(* IEC 61131-3 sources: JingjiangArm/moonboxpro_arm_8.4/Application/Application/数据类型/通讯协议/云影/只写内容/附属内容, 6 files *)

(* ---- StSts_GrpFlag.st ---- *)
(*@CES
Name=StSts_GrpFlag
Type=Gvl
TypeGuid=2db5746d-d284-4425-9f7f-2663a34b0ebc
Guid=84c3180d-bd4c-42e6-a1a9-68017632a9f9
HasDeclaration=True
HasImplementation=False
*)
{DECLARATION}
{attribute 'pack_mode' := '1'}
TYPE StSts_GrpFlag :(*2025.7.3.175755总16字节+8预留字节*)
STRUCT
	xCutterOnTop_Uw								: BIT;(* TRUE=放料上裁 *)
	xCutterOnTop_Rw								: BIT;(* TRUE=放料上裁 *)
	xFlag_Stop									: BIT;(* 停机标志/第1次从当前速度降到空转速度，抬所有色组胶辊/牵引速度到0时抬牵引胶辊，第2次按下则将色组从空转停到0速度 *)
	xFlag_PreStart								: BIT;(* 预启动标志/从停机状态按(预)启动置位标志 色组速度达到空转速度清xFlag_PreStart标志,置位xFlag_Ink标志;当xFlag_Print标志有效后 *)
	xFlag_Ink									: BIT;(* 匀墨标志/>20m/min不能联动 *)
	xFlag_InkAccing								: BIT;(* 匀墨加速中<指0~10m/min那个加速过程> *)
	xFlag_Tension								: BIT;(* 张力投入标志/张力投入有效时收放料变频开始起作用/收放料就位后按印刷按钮,牵引压辊合压/xFlag_Print有效时张力投入不处理 *)
	xFlag_TensionDone							: BIT;(* 张力ok，可以投入印刷 *)
	xFlag_Print									: BIT;(* 张力拉料标志有效时，按联动或印刷按钮 先压收牵(延时2s)再压放牵 印刷标志/印刷色组根据联动标志按用户指定的压辊顺序逐一延时压胶辊/胶辊压合完毕后才可置该标志有效 *)
	xFlag_Estop									: BIT;(* 急停标志/和停机一样要减速到0，只不过减速时间是急停时间 *)
	xFlag_AutoAcc								: BIT;(* 自动加速 *)
	xFlag_AutoDec								: BIT;(* 自动减速 *)
	xFlag_ManuAcc								: BIT;(* 手动加速 *)
	xFlag_ManuDec								: BIT;(* 手动减速 *)
	xFlag_Accing								: BIT;(* 加速中 *)
	xFlag_Decing								: BIT;(* 减速中 *)
	xFlag_EStoping								: BIT;(* 正在急停中 *)
	xFlag_Stoping								: BIT;(* 停机中 *)
	xFlag_GotoInking							: BIT;(* 转到匀墨 *)
	xFlag_InPressing							: BIT;(* 顺序压辊中 *)
	xFlag_RollerPressDone						: BIT;(* 压辊处理完成 *)
	xFlag_InchRun								: BIT;(* 至少有1色处于单运行 *)
	xFlag_AllInchRun							: BIT;(* 整机单运行标志 *)
	xFlag_AllPress								: BIT;(* 全体合压 *)
	xFlag_AllUnpress							: BIT;(* 全体离压 *)
	xFlag_RollerPressAtLeast1					: BIT;(* 至少1色色组合压 *)
	xFlag_PrnLen_Alarm_A						: BIT;
	xFlag_PrnLen_Alarm_B						: BIT;
	xFlag_PrnLen_Alarm_All						: BIT;
	xFlag_LinkageAxisAlarm						: BIT;(* 至少有1个联动轴发生报警 *)
	xFlag_TensionUnfinished						: BIT;(* 张力未完成 *)
	xFlag_VelTooHigh							: BIT;(* 速度过高 *)
	xFlag_PrestartTimeout						: BIT;(* 预启动超时标志 *)
	xFlag_KeepAlarming							: BIT;(* 维持报警*)
	xFlag_ArrivedToTargetVel					: BIT;(* 到达目标速度 *)
	xFlag_FilmAccDecDone						: BIT;(* 料膜加减速完成 *)
	xFlag_IfOf_Ink								: BIT;(*空转牵引联动标志*)
	xFlag_FastStoping							: BIT;
	xSlowStopTenEn								: BIT;(* 收放料慢速松料使能/TRUE *)
	xIsDebugMode_Machine						: BIT;(* 机器调试模式 *)
(*以上40bit*)
	xReflectSensorLoss_Uw						: BIT;(* 放料弧面信号丢失标志/FALSE *)
	xFilmTouchRoller_Uw							: BIT;(*料膜接触到了辊子标志*)
	xSts_PreCutting_Uw							: BIT;(* 放料预备接料/FALSE *)
	xCutterOnTopFroDebug_Uw						: BIT;(* 放料上裁刀标志/用于调试/FALSE *)
	xCurAxisAFroDebug_Uw						: BIT;(* 放料预驱轴为A轴标志/用于调试/FALSE *)
	xAlarmBell_Uw								: BIT;(* 放料响铃常输出/用于控制定位写入响铃提示使用/FALSE *)
	xIsDebuging_DiaMeasure_Uw					: BIT;(* 放料卷径测量调试中/FALSE *)
	xCancelDebuging_DiaMeasure_Uw				: BIT;(* 放料取消卷径测量调试中/FALSE *)
	xEnCodeErr_Uw								: BIT;(* 放料编码器故障*)
	xEnCodeErr_Rw								: BIT;(* 收料编码器故障*)
	xAxisAForeward_Uw							: BIT;(* 放料A轴正转/FALSE *)
	xAxisBForeward_Uw							: BIT;(* 放料B轴正转/FALSE *)
	xFlag_DiamCalc_ing_Uw						: BIT;(* 放料卷径计算中 *)
	xFlag_DiamCalc_end_Uw						: BIT;(* 放料卷径计算完成 *)
	xFlag_DiamMeasure_end_Uw					: BIT;(* 放料卷径测量完成 *)
	xFlag_PreDrv_ing_Uw							: BIT;(* 放料预驱中... *)
	xFlag_PreDrv_end_Uw							: BIT;(* 放料预驱完成  *)
	xFlag_Cut_ing_Uw							: BIT;
	xFlag_Cut_end_Uw							: BIT;
	xFlag_VolDiamAlarm_Uw						: BIT;(* 卷径报警标志 *)
	xStationOnline_AxisA_Uw						: BIT;(* 放料a轴驱动器在线标志/2021.12.4.175524/hdp *)
	xStationOnline_AxisB_Uw						: BIT;(* 放料a轴驱动器在线标志/2021.12.4.175524/hdp *)
	xFlag_AutoMaticCutting_Uw					: BIT;(*2022.4.25.090246 自动裁切中标志*)
(*以上23bit*)
	xSts_PreCutting_Rw							: BIT;(* 收料预备接料 *)
	xCutterOnTopFroDebug_Rw						: BIT;(* 收料上裁刀标志/用于调试/FALSE *)
	xCurAxisAFroDebug_Rw						: BIT;(* 收料预驱轴为A轴标志/用于调试/FALSE *)
	x6InchFroDebug_Rw       					: BIT;(* 收料6寸标志/用于调试/FALSE*)
	xAlarmBell_Rw								: BIT;(* 收料响铃常输出/用于控制定位写入响铃提示使用/FALSE *)
	xAxisAForeward_Rw							: BIT;(* 收料A轴正转/FALSE *)
	xAxisBForeward_Rw							: BIT;(* 收料B轴正转/FALSE *)
	xFlag_6Inch_Rw								: BIT;(* 收料6寸标志/反之为3寸/FALSE *)
	xFlag_PreDrv_ing_Rw							: BIT;(* 收料预驱中... *)
	xFlag_PreDrv_end_Rw							: BIT;(* 收料预驱完成 *)
	xFlag_Cut_ing_Rw							: BIT;(* 收料裁切中 *)
	xFlag_Cut_end_Rw							: BIT;(* 收料裁切完成 *)
	xStationOnline_AxisA_Rw						: BIT;(* 收料a轴驱动器在线标志/2021.12.4.175524/hdp *)
	xStationOnline_AxisB_Rw						: BIT;(* 收料a轴驱动器在线标志/2021.12.4.175524/hdp *)
	xFlag_AutoMaticCutting_rw					: BIT;(*2022.4.25.090246 自动裁切中标志*)
(*以上15bit*)
	xStationOnline_If							: BIT;(* 放牵驱动器在线标志/2021.12.4.175524/hdp *)
	xRollerSts_If								: BIT;(* 放牵压辊/FALSE *)
	xRunEn_If									: BIT;(* 放牵运动使能/0/2021.11.18.201925 *)
	xInching_If									: BIT;(* 放牵单运行中/FALSE *)
	xStationOnline_Of							: BIT;(* 放牵驱动器在线标志/2021.12.4.175524/hdp *)
	xRollerSts_Of								: BIT;(* 放牵压辊/FALSE *)
	xRunEn_Of									: BIT;(* 放牵运动使能/0/2021.11.18.201925 *)
	xInching_Of									: BIT;(* 放牵单运行中/FALSE *)
(*以上8bit*)
	xSts_HorzPreRegister						: BIT;(*横向预套准状态*)
	xFlag_HorzPreRegister_All_end				: BIT;(*横向预套准全部完成*)
	xFlag_Home									: BIT;
	xFlag_Home_ing								: BIT;
	xFlag_Home_end								: BIT;
	xFlag_ConfirmPreRegHomePos					: BIT;(*2017-09-13 12:51:52| 确认预套准基准点*)
	xFlag_ConfirmPreRegHomePos_ing				: BIT;(*确认预套准基准点-ing*)
	xFlag_ConfirmPreRegHomePos_end				: BIT;(*确认预套准基准点-end*)
	xFlag_PreRegister							: BIT;
	xFlag_PreRegister_ing						: BIT;
	xFlag_PreRegister_end						: BIT;
	xFlag_PhaseRestore							: BIT;(*相位恢复*)
	xFlag_PhaseRestore_ing						: BIT;(*相位恢复-ing*)
	xFlag_PhaseRestore_end						: BIT;(*相位恢复-end*)
(*以上14bit*)
	xNetOffline_CENTRAL							: BIT;
	xAxisAlarm_CENTRAL							: BIT;
	xPosDeviationAlarm_CENTRAL					: BIT;
	xNetOffline_CENTRAL2						: BIT;
	xAxisAlarm_CENTRAL2							: BIT;
	xPosDeviationAlarm_CENTRAL2					: BIT;
	xNetOffline_IF								: BIT;
	xAxisAlarm_IF								: BIT;
	xPosDeviationAlarm_IF						: BIT;
	xNetOffline_OF								: BIT;
	xAxisAlarm_OF								: BIT;
	xPosDeviationAlarm_OF						: BIT;
	xNetOffline_UW_A							: BIT;
	xAxisAlarm_UW_A								: BIT;
	xPosDeviationAlarm_UW_A						: BIT;
	xNetOffline_UW_B							: BIT;
	xAxisAlarm_UW_B								: BIT;
	xPosDeviationAlarm_UW_B						: BIT;
	xNetOffline_RW_A							: BIT;
	xAxisAlarm_RW_A								: BIT;
	xPosDeviationAlarm_RW_A						: BIT;
	xNetOffline_RW_B							: BIT;
	xAxisAlarm_RW_B								: BIT;
	xPosDeviationAlarm_RW_B						: BIT;
	xPrintInching								: BIT;//整机点动
	xTapPosition_Breaking						: BIT;(*断料档位|*)
	xTapPosition_UniformInk						: BIT;(*匀墨档位|*)
	xTapPosition_Printing						: BIT;(*印刷档位|*)
(*以上28bit*)
////////////////////////////////////////////////////////////////////////////////////
(*截至这里，以上总共40+23+15+8+14+28=128BIT，占16BYTES，下面再预留8BYTE，用于放系只写标志*)
(*2025.9.18.134744||伪随机中标志-占用一个位预留|niu.j*)
	xPseudoRandomTsting								: BIT;
	xFlag_PressDn_If								: BIT;
	xFlag_PressDn_Of								: BIT;
	xLinkage_If									: BIT;
	xLinkage_Of									: BIT;
//2025.11.14.151756|收放料调试中标bit5\bit6\bit7|新加一个BYTE继续用了bit0||7-1=6
	xFlag_AxisA_DebugRunning_Uw					: BIT;
	xFlag_AxisB_DebugRunning_Uw					: BIT;
	xFlag_AxisA_DebugRunning_Rw					: BIT;
	xFlag_AxisB_DebugRunning_Rw					: BIT;
//	xFlag_GrpRsv5								: BIT;
//	xFlag_GrpRsv6								: BIT;
//	xFlag_GrpRsv7								: BIT;

	xFlag_GrpRsv1								: BIT;
	xFlag_GrpRsv2								: BIT;
	xFlag_GrpRsv3								: BIT;
	xFlag_GrpRsv4								: BIT;
	xFlag_GrpRsv5								: BIT;
	xFlag_GrpRsv6								: BIT;
	xFlag_GrpRsv7								: BIT;

	abyFlag_GrpRsv								: ARRAY [1..6] OF BYTE;
END_STRUCT
END_TYPE

{IMPLEMENTATION}

(* ---- StSts_Modbus.st ---- *)
(*@CES
Name=StSts_Modbus
Type=Gvl
TypeGuid=2db5746d-d284-4425-9f7f-2663a34b0ebc
Guid=cd32acf0-34b3-49da-a704-86f77df9a440
HasDeclaration=True
HasImplementation=False
*)
{DECLARATION}
{attribute 'pack_mode' := '1'}
TYPE StSts_Modbus :
STRUCT
	xCommEn_Tcp								: BIT;(*厂家支持设备tcp通讯使能@常有效*)
	xOpenSocketing							: BIT;(*厂家支持设备tcp打开中@连接中*)
	xOpenSocketDne							: BIT;(*厂家支持设备tcp打开成功*)
	xOpenSocketFailed						: BIT;(*厂家支持设备tcp打开失败*)
	xConnectOk_Tcp							: BIT;(*厂家支持设备连接成功了*)

	(*[1]=监控设备@10bytes*)
	xCommEn_WatchDevice_Tcp					: BIT;(*监控设备tcp通讯使能@常有效*)
	xOpenSocketing_WatchDevice				: BIT;(*监控设备tcp打开中@连接中*)
	xOpenSocketDne_WatchDevice				: BIT;(*监控设备tcp打开成功*)
	xOpenSocketFailed_WatchDevice			: BIT;(*监控设备tcp打开失败*)
	xConnectOk_WatchDevice_Tcp				: BIT;(*监控设备连接成功了*)

(*新增2023.10.14.104239||11字节*)
	(*485需要的@10bytes*)
	xCommEn_485								: BIT;(*485通讯使能开关*)
	xOpenPortDne							: BIT;(*485打开成功*)
	xOpenPortFailed							: BIT;(*485打开失败*)
	xCommEn_WatchDevice_485					: BIT;(*监控设备通讯使能*)

	xRsv_SysFlag_Modbus1					: BIT;(*预留1*)
	xRsv_SysFlag_Modbus2					: BIT;(*预留2*)

	byConnectSts_Tcp						: BYTE;(*厂家支持设备的连接状态		  @=0 未打开
														  @=1 打开中@连接中
														  @=2 打开成功
														  @=3 打开失败
														  @=4 通讯超时*)
	byConnectSts_WatchDevice_Tcp			: BYTE;(*监控设备的连接状态@=0 未打开
														  @=1 打开中@连接中
														  @=2 打开成功
														  @=3 打开失败
														  @=4 通讯超时*)
	byConnectSts_485						: BYTE;(*485设备的连接状态@=0 未打开
											 @=1 打开中@连接中@485不用
											 @=2 打开成功
											 @=3 打开失败*)
	byRsv_SysFlag_Modbus					: BYTE;
END_STRUCT
END_TYPE

{IMPLEMENTATION}

(* ---- StSts_PressRoller_Flag.st ---- *)
(*@CES
Name=StSts_PressRoller_Flag
Type=Gvl
TypeGuid=2db5746d-d284-4425-9f7f-2663a34b0ebc
Guid=b94585e0-0f14-4a6e-b8de-4e371f1e83a5
HasDeclaration=True
HasImplementation=False
*)
{DECLARATION}
{attribute 'pack_mode' := '1'}
TYPE StSts_PressRoller_Flag :(*2025.7.3.175755总2字节+2预留字节*)
STRUCT
	xConfirmAbsEncZeroPosDne_PrnRoller_Pressure_M		: BIT;(* 版辊压力电机绝对值位置M侧/零位确认完成 *)
	xConfirmAbsEncZeroPosDne_PrnRoller_Pressure_G		: BIT;(* 版辊压力电机绝对值位置G侧/零位确认完成 *)
	xConfirmAbsEncZeroPosDne_NetRoller_Pressure_M		: BIT;(* 网辊压力电机绝对值位置M侧/零位确认完成 *)
	xConfirmAbsEncZeroPosDne_NetRoller_Pressure_G		: BIT;(* 网辊压力电机绝对值位置G侧/零位确认完成 *)

(* 2021.12.29.140315/hdp/lyt *)
	xConfirmload_unloadPosDne_PrnRoller_Pressure_M		: BIT;(* 版辊压力电机换版位置M侧/确认完成 *)
	xConfirmload_unloadPosDne_PrnRoller_Pressure_G		: BIT;(* 版辊压力电机换版位置G侧/确认完成 *)
	xConfirmload_unloadPosDne_NetRoller_Pressure_M		: BIT;(* 网辊压力电机换版位置M侧/确认完成 *)
	xConfirmload_unloadPosDne_NetRoller_Pressure_G		: BIT;(* 网辊压力电机换版位置G侧/确认完成 *)

	xConfirmDnPosDne_PrnRoller_Pressure_M				: BIT;(* 版辊压力电机合压位置M侧/确认完成 *)
	xConfirmDnPosDne_PrnRoller_Pressure_G				: BIT;(* 版辊压力电机合压位置G侧/确认完成 *)
	xConfirmDnPosDne_NetRoller_Pressure_M				: BIT;(* 网辊压力电机合压位置M侧/确认完成 *)
	xConfirmDnPosDne_NetRoller_Pressure_G				: BIT;(* 网辊压力电机合压位置G侧/确认完成 *)

	xConfirmDnPosDne_StrRoller_Pressure_M				: BIT;(* 张带辊压力电机合压位置M侧/确认完成 *)
	xConfirmDnPosDne_StrRoller_Pressure_G				: BIT;(* 张带辊压力电机合压位置G侧/确认完成 *)

	xFlag_Rsv0											: BIT;
	xFlag_Rsv1											: BIT;
	abyFlag_Rsv											: ARRAY [1..2] OF BYTE;//预留两个空间
END_STRUCT
END_TYPE

{IMPLEMENTATION}

(* ---- StSts_UnitFlag.st ---- *)
(*@CES
Name=StSts_UnitFlag
Type=Gvl
TypeGuid=2db5746d-d284-4425-9f7f-2663a34b0ebc
Guid=9b5ad9b6-6a41-49ce-aab1-12c5fd79f7c8
HasDeclaration=True
HasImplementation=False
*)
{DECLARATION}
{attribute 'pack_mode' := '1'}
TYPE StSts_UnitFlag :(*2025.7.3.175755总16字节+8预留字节*)
STRUCT
	xLinkage									: BIT;
	xFlag_RollerDn_BottomRoller					: BIT;(* 底辊合压标志/底辊的胶辊 *)
	xFlag_RollerDn_PrnRoller					: BIT;(* 印辊合压标志/靠上底辊 *)
	xFlag_RollerDn_NetRoller					: BIT;(* 网辊合压标志/靠上版辊 *)
	xFlag_HorzPreRegister_ing					: BIT;(*横向预套准进行中|*)
	xFlag_HorzPreRegister_end					: BIT;(*横向预套准完成|*)
	xAxisInching								: BIT;(*版辊单运行中*)
	xAxisInching_Net							: BIT;(*网辊单运行中*)
	xNetOffline_Horz							: BIT;
	xAxisAlarm_Horz								: BIT;
	xPosDeviationAlarm_Horz						: BIT;
	xNetOffline_PrnRoller						: BIT;
	xAxisAlarm_PrnRoller						: BIT;
	xPosDeviationAlarm_PrnRoller				: BIT;
	xNetOffline_NetRoller						: BIT;
	xAxisAlarm_NetRoller						: BIT;
	xPosDeviationAlarm_NetRoller				: BIT;
	xNetOffline_BottomRoller					: BIT;
	xAxisAlarm_BottomRoller						: BIT;
	xPosDeviationAlarm_BottomRoller				: BIT;
	xNetOffline_Prn_Pressure_M					: BIT;
	xAxisAlarm_Prn_Pressure_M					: BIT;
	xPosDeviationAlarm_Prn_Pressure_M			: BIT;
	xNetOffline_Prn_Pressure_G					: BIT;
	xAxisAlarm_Prn_Pressure_G					: BIT;
	xPosDeviationAlarm_Prn_Pressure_G			: BIT;
	xNetOffline_Net_Pressure_M					: BIT;
	xAxisAlarm_Net_Pressure_M					: BIT;
	xPosDeviationAlarm_Net_Pressure_M			: BIT;
	xNetOffline_Net_Pressure_G					: BIT;
	xAxisAlarm_Net_Pressure_G					: BIT;
	xPosDeviationAlarm_Net_Pressure_G			: BIT;
	xNetOffline_Str_Pressure_M					: BIT;
	xAxisAlarm_Str_Pressure_M					: BIT;
	xPosDeviationAlarm_Str_Pressure_M			: BIT;
	xNetOffline_Str_Pressure_G					: BIT;
	xAxisAlarm_Str_Pressure_G					: BIT;
	xPosDeviationAlarm_Str_Pressure_G			: BIT;
	xNetOffline_PHOTOCELL						: BIT;
	xAxisAlarm_PHOTOCELL						: BIT;
	xPosDeviationAlarm_PHOTOCELL				: BIT;
	(*以上总41BIT，预留7bit+2字节*)

	xFlag_PressDn									: BIT;
	xFlag_Rsv2									: BIT;
	xFlag_Rsv3									: BIT;
	xFlag_Rsv4									: BIT;
	xFlag_Rsv5									: BIT;
	xFlag_Rsv6									: BIT;
	xFlag_Rsv7									: BIT;
	abyFlag_Rsv									: ARRAY [1..2] OF BYTE;

END_STRUCT
END_TYPE

{IMPLEMENTATION}

(* ---- StSts_UnitParam.st ---- *)
(*@CES
Name=StSts_UnitParam
Type=Gvl
TypeGuid=2db5746d-d284-4425-9f7f-2663a34b0ebc
Guid=8b49756c-4691-49d4-9f32-1d800649b411
HasDeclaration=True
HasImplementation=False
*)
{DECLARATION}
{attribute 'pack_mode' := '1'}
TYPE StSts_UnitParam :(*总440字节-每个色组两个数据包*)
STRUCT
	diPos_press_dn_PrnRoller_Pressure_M					: DINT;(* 合压位置/版辊压力电机M侧/单位:mm *)
	diPos_press_dn_PrnRoller_Pressure_G					: DINT;(* 合压位置/版辊压力电机G侧/单位:mm *)
	diPos_press_up_PrnRoller_Pressure_M					: DINT;(* 离压位置/版辊压力电机M侧/单位:mm/根据当前合压位置实时变化/2021.12.29.140151 *)
	diPos_press_up_PrnRoller_Pressure_G					: DINT;(* 离压位置/版辊压力电机G侧/单位:mm/根据当前合压位置实时变化/2021.12.29.140151 *)
	diPos_load_unload_PrnRoller_Pressure_M				: DINT;(* 装卸辊位置/版辊压力电机M侧/单位:mm *)
	diPos_load_unload_PrnRoller_Pressure_G				: DINT;(* 装卸辊位置/版辊压力电机G侧/单位:mm *)
	diPos_press_dn_NetRoller_Pressure_M					: DINT;(* 合压位置/网辊压力电机M侧/单位:mm *)
	diPos_press_dn_NetRoller_Pressure_G					: DINT;(* 合压位置/网辊压力电机G侧/单位:mm *)
	diPos_press_up_NetRoller_Pressure_M					: DINT;(* 离压位置/网辊压力电机M侧/单位:mm/根据当前合压位置实时变化/2021.12.29.140151 *)
	diPos_press_up_NetRoller_Pressure_G					: DINT;(* 离压位置/网辊压力电机G侧/单位:mm/根据当前合压位置实时变化/2021.12.29.140151 *)
	diPos_load_unload_NetRoller_Pressure_M				: DINT;(* 装卸辊位置/网辊压力电机M侧/单位:mm *)
	diPos_load_unload_NetRoller_Pressure_G				: DINT;(* 装卸辊位置/网辊压力电机G侧/单位:mm *)
	diPos_press_dn_StrRoller_Pressure_M					: DINT;(* 合压位置/网辊压力电机M侧/单位:mm *)
	diPos_press_dn_StrRoller_Pressure_G					: DINT;(* 合压位置/网辊压力电机G侧/单位:mm *)
	diPos_press_up_StrRoller_Pressure_M					: DINT;(* 离压位置/网辊压力电机M侧/单位:mm/根据当前合压位置实时变化/2021.12.29.140151 *)
	diPos_press_up_StrRoller_Pressure_G					: DINT;(* 离压位置/网辊压力电机G侧/单位:mm/根据当前合压位置实时变化/2021.12.29.140151 *)
	diPos_load_unload_StrRoller_Pressure_M				: DINT;(* 装卸辊位置/网辊压力电机M侧/单位:mm *)
	diPos_load_unload_StrRoller_Pressure_G				: DINT;(* 装卸辊位置/网辊压力电机G侧/单位:mm *)
	diGirth_Confirmed_press_dn_PrnRoller				: DINT;(* 确认合压位时候的版辊周长*)
	diGirth_Confirmed_press_dn_NetRoller				: DINT;(* 确认合压位时候的网纹辊周长*)
	diGirth_Confirmed_press_dn_StrRoller				: DINT;(* 确认合压位时候的网纹辊周长*)
	stStSts_PressRoller_Flag							: StSts_PressRoller_Flag;
(*该结构体StSts_PressRoller_Flag----4*MAX_UNIT_NUM字节-64字节*)

	rAI_med_CoatingPrn									: REAL;(*涂布中位值|*)
	(*bit0-bit15分别对应色组1到16*)
	diEncPosPrintDn_Prn_M 								: DINT;
	diEncPosPrintDn_Prn_G 								: DINT;
	diEncPosPrintDn_Net_M 								: DINT;
	diEncPosPrintDn_Net_G 								: DINT;
	diEncPosPrintDn_Str_M 								: DINT;
	diEncPosPrintDn_Str_G 								: DINT;
		//2024.10.21.114530 | bai.zy | 版辊网辊操作侧传动侧平行位置标定值	48字节
	diEncPosParallel_Prn_M 							: DINT;
	diEncPosParallel_Prn_G 							: DINT;
	diEncPosParallel_Net_M 							: DINT;
	diEncPosParallel_Net_G 							: DINT;
	diEncPosParallel_Str_M 							: DINT;
	diEncPosParallel_Str_G 							: DINT;
		//2024.10.21.114530 | bai.zy | 版辊网辊操作侧传动侧合压位偏移量	  48字节
	diPrintPosOffsetDn_Prn_M 							: DINT;
	diPrintPosOffsetDn_Prn_G 							: DINT;
	diPrintPosOffsetDn_Net_M 							: DINT;
	diPrintPosOffsetDn_Net_G 							: DINT;
	diPrintPosOffsetDn_Str_M 							: DINT;
	diPrintPosOffsetDn_Str_G 							: DINT;
	diSampleNum 										: DINT;//采样减速比分子
	diSampleDen 										: DINT;//采样减速比分母
	rSampleGirth										: REAL;
//2024.11.27.154753 | bai.zy | 增加绝对编码器位置,48字节
	diABSPos_Prn_M										: DINT;
	diABSPos_Prn_G 									: DINT;
	diABSPos_Net_M 									: DINT;
	diABSPos_Net_G 									: DINT;
	diABSPos_Str_M 									: DINT;
	diABSPos_Str_G 									: DINT;

	diEncPosLimit_Prn_M_Max 							: DINT;
	diEncPosLimit_Prn_G_Max 							: DINT;
	diEncPosLimit_Net_M_Max 							: DINT;
	diEncPosLimit_Net_G_Max 							: DINT;
	diEncPosLimit_Str_M_Max 							: DINT;
	diEncPosLimit_Str_G_Max 							: DINT;
	rPos_press_dn_PrnRoller_Pressure_M_Hmi				: REAL;(* 根据坐标系界面显示变量-hmi/合压位置/版辊压力电机M侧/单位:mm *)
	rPos_press_dn_PrnRoller_Pressure_G_Hmi				: REAL;(* 根据坐标系界面显示变量-hmi/合压位置/版辊压力电机G侧/单位:mm *)
	rPos_press_up_PrnRoller_Pressure_M_Hmi				: REAL;(* 根据坐标系界面显示变量-hmi/离压位置/版辊压力电机M侧/单位:mm *)
	rPos_press_up_PrnRoller_Pressure_G_Hmi				: REAL;(* 根据坐标系界面显示变量-hmi/离压位置/版辊压力电机G侧/单位:mm *)
	rPos_load_unload_PrnRoller_Pressure_M_Hmi			: REAL;(* 根据坐标系界面显示变量-hmi/装卸辊位置/版辊压力电机M侧/单位:mm *)
	rPos_load_unload_PrnRoller_Pressure_G_Hmi			: REAL;(* 根据坐标系界面显示变量-hmi/装卸辊位置/版辊压力电机G侧/单位:mm *)
	rPos_press_dn_NetRoller_Pressure_M_Hmi				: REAL;(* 根据坐标系界面显示变量-hmi/合压位置/网辊压力电机M侧/单位:mm *)
	rPos_press_dn_NetRoller_Pressure_G_Hmi				: REAL;(* 根据坐标系界面显示变量-hmi/合压位置/网辊压力电机G侧/单位:mm *)
	rPos_press_up_NetRoller_Pressure_M_Hmi				: REAL;(* 根据坐标系界面显示变量-hmi/离压位置/网辊压力电机M侧/单位:mm *)
	rPos_press_up_NetRoller_Pressure_G_Hmi				: REAL;(* 根据坐标系界面显示变量-hmi/离压位置/网辊压力电机G侧/单位:mm *)
	rPos_load_unload_NetRoller_Pressure_M_Hmi			: REAL;(* 根据坐标系界面显示变量-hmi/装卸辊位置/网辊压力电机M侧/单位:mm *)
	rPos_load_unload_NetRoller_Pressure_G_Hmi			: REAL;(* 根据坐标系界面显示变量-hmi/装卸辊位置/网辊压力电机G侧/单位:mm *)
	rPos_PrnRoller_Pressure_M							: REAL;(* 版辊压力电机位置M侧/实时值|mm-根据坐标系变化 *)
	rPos_PrnRoller_Pressure_G							: REAL;(* 版辊压力电机位置G侧/实时值|mm-根据坐标系变化 *)
	rPos_NetRoller_Pressure_M							: REAL;(* 网辊压力电机位置M侧/实时值|mm-根据坐标系变化 *)
	rPos_NetRoller_Pressure_G							: REAL;(* 网辊压力电机位置G侧/实时值|mm-根据坐标系变化 *)
	rPos_StrRoller_Pressure_M							: REAL;(* 张带辊压力电机位置M侧/实时值|mm-根据坐标系变化 *)
	rPos_StrRoller_Pressure_G							: REAL;(* 张带辊压力电机位置G侧/实时值|mm-根据坐标系变化 *)
	dwAxisAlrSts_NetRoller_Pressure_M					: DWORD;(* 网辊压力M侧报警状态 *)
	dwAlrCode_NetRoller_Pressure_M						: DWORD;(* 网辊压力M侧报警代码 *)
	dwAxisAlrSts_NetRoller_Pressure_G					: DWORD;(* 网辊压力G侧报警状态 *)
	dwAlrCode_NetRoller_Pressure_G						: DWORD;(* 网辊压力G侧报警代码 *)
	dwAxisAlrSts_PrnRoller_Pressure_M					: DWORD;(* 版辊压力M侧报警状态 *)
	dwAlrCode_PrnRoller_Pressure_M						: DWORD;(* 版辊压力M侧报警代码 *)
	dwAxisAlrSts_PrnRoller_Pressure_G					: DWORD;(* 版辊压力G侧报警状态 *)
	dwAlrCode_PrnRoller_Pressure_G						: DWORD;(* 版辊压力G侧报警代码 *)
	dwAlarmDetail_Prn									: DWORD;//轴报警信息-版辊
	dwAlarmDetail_Net									: DWORD;//轴报警信息-wnag辊
	dwAlarmDetail_Bottom								: DWORD;//轴报警信息-底辊
	dwAlarmDetail_Prn_M								: DWORD;//轴报警信息-版辊_M
	dwAlarmDetail_Prn_G								: DWORD;//轴报警信息-版辊_G
	dwAlarmDetail_Net_M								: DWORD;//轴报警信息-网辊_M
	dwAlarmDetail_Net_G								: DWORD;//轴报警信息-网辊_G
	dwAlarmDetail_Horz									: DWORD;//轴报警信息-横向
	dwAlarmDetail_PHOTOCELL							: DWORD;//光电眼
	dwAlarmDetail_Str_M								: DWORD;//轴报警信息-网辊_M
	dwAlarmDetail_Str_G								: DWORD;//轴报警信息-网辊_G
	rPhotoCellPosLimit_M 								: REAL;
	rPhotoCellPosLimit_G 								: REAL;

(*该结构体8字节*MAX_UNIT_NUM=128字节*)
	stStSts_UnitFlag									: StSts_UnitFlag;

	rPV_UnitTemCtl										: REAL;(* 色组温度控制实时值 *)
	rHz_UnitExhaust_CurrRD								: REAL;(* 排风当前回读频率/pdu上行给主站/ *)
	rHz_UnitExhaust_CurrWR								: REAL;(* 排风当前写入频率/pdu下行给从站/ *)
	rHz_UnitHotWind2_CurrRD							: REAL;(* 热风当前回读频率/pdu上行给主站/ *)
	rHz_UnitHotWind2_CurrWR							: REAL;(* 热风当前写入频率/pdu下行给从站/ *)
	rHz_UnitHotWind_CurrRD								: REAL;(* 热风当前回读频率/pdu上行给主站/ *)
	rHz_UnitHotWind_CurrWR								: REAL;(* 热风当前写入频率/pdu下行给从站/ *)
	rHz_UnitScraper_CurrRD								: REAL;(* 刮刀当前回读频率/pdu上行给主站/ *)
	rHz_UnitScraper_CurrWR								: REAL;(* 刮刀当前写入频率/pdu下行给从站/ *)
	rHz_UnitInkRoller_CurrRD							: REAL;(* 递墨辊当前回读频率/pdu上行给主站/ *)
	rHz_UnitInkRoller_CurrWR							: REAL;(* 递墨辊当前写入频率/pdu下行给从站/ *)

(*	//增加色组版辊相位2025.8.25.152919					|niu.j*)
	wVirtual											: WORD;
//2025.10.20.151557增加预套准料长值||6-4=2
	rPreReg_Length_V						: REAL;(*纵向预套准料长值|单位:mm|*)
//增加色组版辊虚拟码盘状态--2字节
	wVirTual_Sts										: WORD;
//	abyRsv												: ARRAY [1..2] OF BYTE;
END_STRUCT
END_TYPE
{IMPLEMENTATION}

(* ---- StSts_UnitParam_2.st ---- *)
(*@CES
Name=StSts_UnitParam_2
Type=Gvl
TypeGuid=2db5746d-d284-4425-9f7f-2663a34b0ebc
Guid=204de66d-e1be-420b-af3f-8c8766064217
HasDeclaration=True
HasImplementation=False
*)
{DECLARATION}
{attribute 'pack_mode' := '1'}
TYPE StSts_UnitParam_2 :(*总110字节，两个色组一个数据包*)(*2025.7.3.175755增加330字节预留-总440字节*)
STRUCT

	byCurPos_Roller									: BYTE;(*辊子当前位置|0 换版位
																		  1 离压位
																		  2 合压位*)
	byInPos_Roller										: BYTE;(*辊子到位标志|.0 全部到位
																		  .1 版辊操作侧到位
																		  .2 版辊传动侧到位
																		  .3 网辊操作侧到位
																		  .4 网辊传动侧到位*)
	byColorIdCurrent									: BYTE;(*当前色序				*)
	byColorIdFollow									: BYTE;(*跟踪色序				*)
	byArcSts											: BYTE;(* 套色状态/bit0=报警/bit1=丢失 *)
	wSts_HorzManuPreReg								: WORD; (* 横向手动预套准状态标志|bit0运行标志|bit1正转|bit2反转|bit3左限位|bit4右限位|bit5停止 *)
	iPos_HorzManuPreReg								: INT;(*横向手动预套准位置|*)
	wSTS_UnitExhaust									: WORD;(* 排风状态|/.0 通讯返回运行状态
															   /.6 排风打开超时-
															   /.7 485通讯断开标志
															   高8位作为报警码*)
(*	原来的接口，先不要了				作为预留6字节
	wUnit_input_I 										: WORD;
	wUnit_input_II 									: WORD;
	wUnit_input_III 									: WORD;
	*)

//2025.12.30.223243增加风门当前位置显示||6-4=2
	rUnitExhaustDamperPos_Cur				: REAL;(*排风风门写入当前位置值*)
	abyRsv_Data_1										: ARRAY [1..2] OF BYTE;

	wSTS_UnitHotWind_2									: WORD;(* 热风II状态 *)
	wSTS_UnitHotWind									: WORD;(* 热风状态 |.0 运行\停止
															               /.6 热风风打开超时-
															  			   /.7 485通讯断开标志*)
	wSTS_UnitScraper									: WORD;(* 刮刀状态/pdu上行给主站/ |.0 运行\停止
															              				  /.6 刮刀打开超时-
															                              /.7 485通讯断开标志*)
	wSTS_UnitInkRoller									: WORD;(* 递墨辊状态/pdu上行给主站 |.0 运行\停止
															              				   /.6 递墨辊刀打开超时
															                               /.7 485通讯断开标志*)
	wSTS_UnitTemCtl									: WORD;(* 色组温度控制报警代码|低8位作为运行状态
																				/.0 通讯返回运行状态
																				/.1 加热使能输出状态
												  高8位作为报警状态/.8 断偶标志
																   /.9 超温标志
																   /.10 离线标志*)

	awInput_IOTestDI_Axis							: ARRAY [1..7] OF WORD;
	awInput_IOTestDI_Axis_Extra						: ARRAY [1..7] OF WORD;
	awInput_IOTestAI_Axis							: ARRAY [1..6] OF WORD;
	awInput_IOTestAI_Axis_Extra						: ARRAY [1..16] OF WORD;
(*增加IO监控2025.8.20.153450*)

//2025.10.15.163922||增加涂布模拟量和轴速度||11-8=3
	rAI_Coating									: REAL;   //涂布摆臂值
	rVel_Coating								: REAL;	//涂布轴速度

//增加一些秦华相关的2025.12.31.112154||总共14字节||113-14=99
	rLength_Band								: REAL;//带长
	iTriggerCnt									: INT;//DI触发
	udiTriggerTimeErr							: UDINT;//DI时间
	udiTriggerEncErr							: UDINT;//DI编码器
//2026.2.2.160436||增加柔印相关一些内容；||niu.j||总12字节99-12= 87；
	rParallelError_Prn_MM						: REAL;
	rParallelError_Net_MM						: REAL;
	rParallelError_Str_MM						: REAL;
//2026.4.25.141239增加全自动套印相关内容2026.4.25.141251
//6字节
	wCommFromDubheFindSignal 	: WORD;//:WORD;(*Bit0 xFlag_AutoAdj_En:BOOL;(*该轴全自动套印使能*)
										//Bit1 xFlag_FindFirstSuccess					: BOOL;(*找到当前色完成*)
										//Bit2 xFlag_FindPreSuccess					: BOOL;(*找到前一色*)
										//Bit3 xFlag_AutoAdj_En:BOOL;(*该轴全自动套印完成*)			）
										//Bit4 xCurManuAdjust :BOOL;(*当前色未找到，需要手动调整光电眼位置，调整好后人工置位*)-----------------Reset
										//Bit5 xPreCurManuAdjust :BOOL;(*前一色未找到，需要观察原因调整好后，人工点确定，等一个机组料长后置位*)
										//*)
	iError_Msg					: INT;//	: INT;(*0:无错误                 -------------------------------------------错误码
										//-1~-100:单色色标失败原因
										//-101~-200:混色色标失败原因*)
	iStep_AutoAdjust 			: INT;//:  INT;(*主站全自动套印的找标的执行状态   -------------------步骤码*)

//结束2026.4.25.141327

//2026.4.25.142714部分两个变量不需要双向通讯|2变量8字节|81-8=73
	rKp_MolCal                     					: REAL;
	rKi_MolCal                     					: REAL;

//2026.06.15.184209 增加电压实时值0-220v 增加电压实时值0-220v 73-3=70
	abyVoltage_PV:ARRAY [1..3] OF BYTE;

//2026.06.29.200311||增加横向伺服当前位置单向只写70-4=66
	diPos_Horz									:DINT;

	abyDataRsv										: ARRAY [1..66] OF BYTE;

//////////////////////////////////////分界线-每隔一段数据增加些预留空间/////////////////////////////////////////////////////////////////////////////
	abyRsvData_c										: ARRAY [1..220] OF BYTE;
//////////////////////////////////////////////////////////////////////////////////////////////////////////////////////////////////////////
END_STRUCT
END_TYPE

{IMPLEMENTATION}
